// TIA Portal V20 export
DATA_BLOCK "POS3_0_Melden_Visu_DB"   // DB62
// stored: AssignedProDiagFB POS3_0_Prodiag, InstanceOfName POS3_0_Melden_Visu, InstanceOfType FB
"POS3_0_Melden_Visu"
   // VAR
   //    "Taktzeitermittlung_mit_WT-Wechsel" { S7_SetPoint := 'True'} : "Taktzeitermittlung_Start_Stop_V1_0";
   //    Taktzeitermittlung { S7_SetPoint := 'True'} : "Taktzeitermittlung_Start_Stop_V1_0";
   //    R_TRIG_Init_Achse_1 { S7_SetPoint := 'True'} : R_TRIG;
   //    R_TRIG_Init_Achse_1_Positionen { S7_SetPoint := 'True'} : R_TRIG;
   //    R_TRIG_Init_Achse_2 { S7_SetPoint := 'True'} : R_TRIG;
   //    R_TRIG_Init_Achse_2_Positionen { S7_SetPoint := 'True'} : R_TRIG;
   //    Zyklen_für_Durchschnittszeit { ExternalAccessible := 'False'; ExternalVisible := 'False'; ExternalWritable := 'False'} : Int;
   //    Summe { ExternalAccessible := 'False'; ExternalVisible := 'False'; ExternalWritable := 'False'} : Real;
   // END_VAR
BEGIN
END_DATA_BLOCK
